Fanuc KAREL source: ko00091.KL

-- PROVISIONAL review KL for V1013-1; original PC SHA256 39d1cd9533f9ab2e6500538b46ff485035f54361c340d59ae6148cd26c9891d6
-- Incomplete behavior may be omitted. Consult companion uncertainty JSON. Do not deploy.
PROGRAM KO00091
%NOLOCKGROUP
BEGIN
  -- UNRESOLVED_PC offsets 5-12; opcodes 9D,23
  -- UNRESOLVED_PC offsets 17-69; opcodes 27,27,49,7E,AD,27,49,7E,AD,22,31,7E,4A
  -- UNRESOLVED_PC offsets 74-78; opcodes 7F
END KO00091
